Staubli VAL3: HMI_cs9.pjx

--- HMI_cs9.pjx ---
Parameters version=s8.10.3Cs9_BS2093 stackSize=5000 millimeterUnit=true
Program file=main.pgx
Program file=start.pgx
Program file=stop.pgx
Data file=HMI_cs9.dtx
Library alias=rs path=Disk://source/projectSource/robotStatus/robotStatus.pjx
Library alias=util path=./HMI_util/HMI_util.pjx
Library alias=io path=./HMI_action/HMI_action.pjx
Library alias=home path=./home/home.pjx

--- HMI_cs9.dtx ---
mdesc mNomSpeed

--- main.pgx ---
public program main()
begin
  if rs:sPageUsing!="main"
    rs:sPageUsing="main"
    //
    call util:loadingPage()
    //
    userPage(rs:sPageUsing)
    delay(1)
  endIf
end

--- start.pgx ---
program start()
begin
  call home:main()
end

--- stop.pgx ---
program stop()
begin
end
